FUNCTION_BLOCK ALARM_RING (* Migrated from IEC 61131-3 ST *)
  (* Standard: 61499-2 *)
  (* Version 1.0, 2026-11-06, st2fb *)
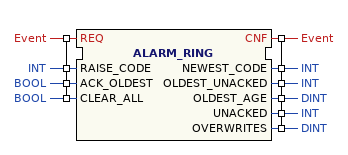
  EVENT_INPUT
    REQ WITH RAISE_CODE, ACK_OLDEST, CLEAR_ALL;
  END_EVENT
  EVENT_OUTPUT
    CNF WITH NEWEST_CODE, OLDEST_UNACKED, OLDEST_AGE, UNACKED, OVERWRITES;
  END_EVENT
  VAR_INPUT
    RAISE_CODE : INT;
    ACK_OLDEST : BOOL;
    CLEAR_ALL : BOOL;
  END_VAR
  VAR_OUTPUT
    NEWEST_CODE : INT;
    OLDEST_UNACKED : INT;
    OLDEST_AGE : DINT;
    UNACKED : INT;
    OVERWRITES : DINT;
  END_VAR
  VAR
    RING_CODE_1 : INT := 0;
    RING_CODE_2 : INT := 0;
    RING_CODE_3 : INT := 0;
    RING_CODE_4 : INT := 0;
    RING_ACKED_1 : BOOL := FALSE;
    RING_ACKED_2 : BOOL := FALSE;
    RING_ACKED_3 : BOOL := FALSE;
    RING_ACKED_4 : BOOL := FALSE;
    RING_AGE_1 : DINT := 0;
    RING_AGE_2 : DINT := 0;
    RING_AGE_3 : DINT := 0;
    RING_AGE_4 : DINT := 0;
    HEAD : INT := 1;
    USED : INT := 0;
    I : INT := 0;
    SLOT : INT := 0;
    PREV_CODE : INT := 0;
    ACK_EDGE_CLK : BOOL := FALSE;
    ACK_EDGE_Q : BOOL := FALSE;
    ACK_EDGE_M : BOOL := FALSE;
    FOUND : BOOL := FALSE;
    CUR_CODE : INT := 0;
    CUR_ACKED : BOOL := FALSE;
    CUR_AGE : DINT := 0;
  END_VAR
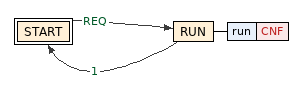
  EC_STATES
    START;
    RUN : run -> CNF;
  END_STATES
  EC_TRANSITIONS
    START TO RUN := REQ;
    RUN TO START := 1;
  END_TRANSITIONS
  ALGORITHM run IN ST:
ACK_EDGE_CLK := ACK_OLDEST;
ACK_EDGE_Q := ACK_EDGE_CLK AND NOT ACK_EDGE_M;
ACK_EDGE_M := ACK_EDGE_CLK;

IF CLEAR_ALL THEN
  RING_CODE_1 := 0; RING_CODE_2 := 0; RING_CODE_3 := 0; RING_CODE_4 := 0;
  RING_ACKED_1 := FALSE; RING_ACKED_2 := FALSE; RING_ACKED_3 := FALSE; RING_ACKED_4 := FALSE;
  RING_AGE_1 := 0; RING_AGE_2 := 0; RING_AGE_3 := 0; RING_AGE_4 := 0;
  HEAD := 1;
  USED := 0;
  NEWEST_CODE := 0;
ELSIF (RAISE_CODE <> 0) AND (RAISE_CODE <> PREV_CODE) THEN
  IF USED = 4 THEN
    OVERWRITES := OVERWRITES + 1;
  ELSE
    USED := USED + 1;
  END_IF;
  CASE HEAD OF
    1: RING_CODE_1 := RAISE_CODE; RING_ACKED_1 := FALSE; RING_AGE_1 := 0;
    2: RING_CODE_2 := RAISE_CODE; RING_ACKED_2 := FALSE; RING_AGE_2 := 0;
    3: RING_CODE_3 := RAISE_CODE; RING_ACKED_3 := FALSE; RING_AGE_3 := 0;
    4: RING_CODE_4 := RAISE_CODE; RING_ACKED_4 := FALSE; RING_AGE_4 := 0;
  END_CASE;
  NEWEST_CODE := RAISE_CODE;
  HEAD := HEAD MOD 4 + 1;
END_IF;
PREV_CODE := RAISE_CODE;

OLDEST_UNACKED := 0;
OLDEST_AGE := 0;
UNACKED := 0;
FOR I := 1 TO USED DO
  SLOT := (HEAD - USED + I + 3) MOD 4 + 1;
  CASE SLOT OF
    1: RING_AGE_1 := RING_AGE_1 + 1;
    2: RING_AGE_2 := RING_AGE_2 + 1;
    3: RING_AGE_3 := RING_AGE_3 + 1;
    4: RING_AGE_4 := RING_AGE_4 + 1;
  END_CASE;
END_FOR;
IF ACK_EDGE_Q THEN
  FOUND := FALSE;
  FOR I := 1 TO USED DO
    IF NOT FOUND THEN
      SLOT := (HEAD - USED + I + 3) MOD 4 + 1;
      CASE SLOT OF
        1: CUR_ACKED := RING_ACKED_1;
        2: CUR_ACKED := RING_ACKED_2;
        3: CUR_ACKED := RING_ACKED_3;
        4: CUR_ACKED := RING_ACKED_4;
      END_CASE;
      IF NOT CUR_ACKED THEN
        CASE SLOT OF
          1: RING_ACKED_1 := TRUE;
          2: RING_ACKED_2 := TRUE;
          3: RING_ACKED_3 := TRUE;
          4: RING_ACKED_4 := TRUE;
        END_CASE;
        FOUND := TRUE;
      END_IF;
    END_IF;
  END_FOR;
END_IF;
FOR I := USED TO 1 BY -1 DO
  SLOT := (HEAD - USED + I + 3) MOD 4 + 1;
  CASE SLOT OF
    1: CUR_ACKED := RING_ACKED_1; CUR_CODE := RING_CODE_1; CUR_AGE := RING_AGE_1;
    2: CUR_ACKED := RING_ACKED_2; CUR_CODE := RING_CODE_2; CUR_AGE := RING_AGE_2;
    3: CUR_ACKED := RING_ACKED_3; CUR_CODE := RING_CODE_3; CUR_AGE := RING_AGE_3;
    4: CUR_ACKED := RING_ACKED_4; CUR_CODE := RING_CODE_4; CUR_AGE := RING_AGE_4;
  END_CASE;
  IF NOT CUR_ACKED THEN
    UNACKED := UNACKED + 1;
    OLDEST_UNACKED := CUR_CODE;
    OLDEST_AGE := CUR_AGE;
  END_IF;
END_FOR;
  END_ALGORITHM
END_FUNCTION_BLOCK
